(* IEC 61131-3 sources: 2026_Projet_YGO_ExcavatriceDragage/CODE_BACKUP/CODE_20260907_ChantierWeekEnd_v0.6.43/G_CYCLE/_TYPES, 10 files *)

(* ---- E_AutoCycleStep.st ---- *)
(* =======================================================================
   ⚙️ E_AutoCycleStep — Etapes du GRAFCET du cycle SEMI_AUTO (dragage)
   ───────────────────────────────────────────────────────────────
   🎯 Role : Enumeration des steps du sequenceur SEMI_AUTO (FB_CycleSemiAuto).
             Prefixe AX (Auto) homogene au homing machine (prefixe HX).
   📄 Doc metier : DOC/AF/AF_Partie-04_Mode_SemiAuto_Sequenceur_v2.3.md
                   + DOC/WFLOW/CONTRACTS/GEL_GRAFCET_SEMIAUTO_20260903.md
   🧊 GEL 2026-09-03 : DIVING decompose en 5 steps de plein droit (AX4..AX8) +
             step special AX_DIVING_RETRY ; EXTRACTION = AX9..AX12 ;
             DECHARGE = AX13..AX15C + AX18_DONE_SYNC ; AX_STAB repli defaut.
   ======================================================================= *)

TYPE E_AutoCycleStep :
(
  AX0_REPOS             := 0,   (* Repos / park : toutes commandes 0, etat neutre - etape initiale pure *)
  AX1_INIT             := 1,    (* Verif CONDITIONS INITIALES (Homed M1/M2, treuils FDC haut, M3 pas a droite de P1) - aucun mouvement, aucun referencement *)
  AX2_TRANSLATE_P1     := 2,    (* Translation vers P1 : joystick vers la droite, le cycle n'emet aucune commande M3 ; surveillance treuils au FDC haut *)
  AX3_OPEN_BUCKET      := 3,    (* Ouverture benne jusqu'au FDC logiciel benne ouverte *)

  (* --- DIVING (5 steps + retry) --- *)
  AX4_DESCEND_DIVING   := 4,    (* Plongee couplee benne ouverte palier 4 jusqu'a l'altimetrie de lancement (DiveStartMin_M) - Kobold PAS enclenche *)
  AX5_KOBOLD_INIT      := 5,    (* Activation contacteur Kobold << au vol >>, verif retour contacteur, descente palier 4 maintenue *)
  AX6_SEARCH_IMMERSION := 6,    (* Recherche entree dans l'eau : attente front DI Kobold 0->1, descente palier 4 maintenue *)
  AX7_SEARCH_BOTTOM    := 7,    (* Recherche du fond : attente front DI Kobold 1->0, descente palier 4 maintenue *)
  AX8_BOTTOM_CONFIRMED := 8,    (* Fond confirme : coupure instantanee treuils, set bit fond, TouchPositionM / RaiseTargetM *)

  (* --- EXTRACTION (4 steps) --- *)
  AX9_RAISE_OFF_BOTTOM := 9,    (* Montee synchronisee : retendre les cables ; selecteur couplage BOTH/M1/M2 accessible *)
  AX10_CLOSE_BUCKET    := 10,   (* Fermeture benne, treuils explicitement 0 *)
  AX11_CTRL_ASCENT     := 11,   (* Montee controle palier max reglable [1..2] + surveillance ecart vitesse M1/M2 ; benne mal fermee autorisee *)
  AX12_LOADED_ASCENT   := 12,   (* Montee en charge : palier 4 si benne fermee, palier 1 si mal fermee ; pas de ralenti 1 m avant top *)

  (* --- DECHARGE (6 steps) --- *)
  AX13_DRAIN_PAUSE     := 13,   (* Egouttage temporise - duree reglable IHM + bypass immediat *)
  AX14_TRANSLATE_DUMP  := 14,   (* Translation vers tremie (depart P1) + avertissements IHM *)
  AX15A_DUMP_ARRIVE    := 15,   (* Arrivee tremie : treuils a l'arret, attente geste operateur *)
  AX15B_DUMP_OPEN      := 16,   (* Vidage : ouverture benne au-dessus de la tremie, LES DEUX treuils a l'arret *)
  AX15C_DUMP_REPOSITION := 17,  (* Repositionnement couple M1+M2 (option IHM maintenue), retour AX15B au relachement *)
  AX18_DONE_SYNC       := 18,   (* Fin de passe : compteur vidages + duree cycle ; msg << aller en P1 >> ; rebouclage direct sur AX2 *)

  (* --- STEPS SPECIAUX --- *)
  AX_STAB              := 19,   (* Repli defaut / stabilisation - pas une erreur *)
  AX_DIVING_RETRY      := 20,   (* Reprise diving : remontee assistee palier lent jusqu'au FDC haut puis retour AX4 ; sur erreur Kobold / joystick relache / palier <> 4 en AX5..AX7 *)
  AX3_WAIT_DIVE_START  := 21,   (* Transition benne->plongee : sorties neutres jusqu'a l'arret mecanique confirme M1/M2, joystick pousse maintenu *)
  AX10_WAIT_ASCENT_START := 22  (* Transition fermeture->montee : sorties neutres jusqu'a l'arret confirme M1/M2, joystick tire maintenu *)
);
END_TYPE

(* ---- E_MachineHomingStep.st ---- *)
(* =======================================================================
   ⚙️ E_MachineHomingStep — Etapes du guide de referencement machine
   ───────────────────────────────────────────────────────────────
   🎯 Rôle : Etat publie du guide de homing conjoint M1/M2/benne (IHM + interlocks)
   📄 Doc métier : DOC/AF/AF_Partie-09_Fonction_Encoder_v2.4.md (F09.08)
   ======================================================================= *)

TYPE E_MachineHomingStep :
(
    IDLE                 := 0,   (* Referencement indisponible (Enable=FALSE) *)
    LOSS_SAFESTOP        := 5,   (* Perte de datum en mouvement : arret controle en cours *)
    BOTH_NOT_HOMED       := 10,  (* Codeurs M1 et M2 non references : passer en MAINT_N2 *)
    M1_NOT_HOMED         := 11,  (* Codeur M1 non reference ou mesure douteuse : homer M1 *)
    M2_NOT_HOMED         := 12,  (* Codeur M2 non reference ou mesure douteuse : homer M2 *)
    OFFSET_UNKNOWN       := 20,  (* Offset benne inconnu : passer en MAINT_N2 *)
    NEED_TOP_POSITION    := 30,  (* Monter Both a vitesse lente jusqu au capteur haut *)
    NEED_MECHANICAL_STOP := 40,  (* Capteur haut atteint : relacher la commande et attendre l arret *)
    AWAIT_BUCKET_CONFIRM := 45,  (* Confirmer visuellement la benne : Fermee ou Ouverte *)
    HOMING_IN_PROGRESS   := 50,  (* Referencement conjoint M1/M2 en cours : ne pas manoeuvrer *)
    VALID                := 60,  (* Referencement machine valide : mode nominal disponible *)
    FAILED               := 70   (* Referencement incomplet : rester en N2 et recommencer *)
);
END_TYPE

(* ---- E_MachineHomingTxState.st ---- *)
(* =======================================================================
   ⚙️ E_MachineHomingTxState — Steps du GRAFCET de referencement machine
   ───────────────────────────────────────────────────────────────
   🎯 Role : Machine a etats sequentielle (GRAFCET) du cycle de homing
             machine M1/M2/benne pilote par FB_CycleMachineHoming (§4).
             Distincte de E_MachineHomingStep (echelle de priorite du
             guide operateur, libelles de diagnostic - §6).
   📄 Doc : DOC/WFLOW/CONTRACTS/GEL_GRAFCET_HOMING_CYCLE_20260903.md
            + DOC/AF/AF_Partie-09_Fonction_Encoder_v2.4.md (F09.08)
   ======================================================================= *)

TYPE E_MachineHomingTxState :
(
    HX0_REPOS         := 0,   (* Etape initiale pure : aucune action, aucune affectation *)
    HX1_CHOICE        := 1,   (* Annonce + choix operateur : aucun mouvement *)
    HX2_CLIMB         := 2,   (* Chemin A : montee couplee M1+M2 palier 1 jusqu au capteur haut *)
    HX2N_NEUTRAL      := 3,   (* Arret + inversion de sens (tire -> pousse) : mouvement nul obligatoire *)
    HX3_HOME_AXES     := 4,   (* Homing axes M1+M2 au vol sur front descendant capteur, puis descente couplee *)
    HX3N_PAUSE        := 5,   (* Arret avant benne : mouvement nul, retour joystick au neutre *)
    HX4_BUCKET_ADJUST := 6,   (* Ajustement benne palier 1 sans FDC soft, 2 sens autorises *)
    HX5_BUCKET_COMMIT := 7,   (* Commit atomique etat benne fermee (CommitClose) *)
    HX6_HOMED         := 8,   (* Machine referencee : MachineHomed := TRUE (fugace) *)
    HXF_FAILED        := 9    (* Referencement incomplet : rester en N2 et recommencer *)
);
END_TYPE

(* ---- E_OperatorAxis.st ---- *)
(* =======================================================================
   ⚙️ E_OperatorAxis — Axe ou organe de pilotage attendu par le cycle
   ───────────────────────────────────────────────────────────────
   🎯 Rôle : Énumération de l'organe joystick/bouton attendu pour le mouvement
   📄 Doc métier : DOC/AF/AF_Partie-04_Mode_SemiAuto_Sequenceur_v2.3.md
   ======================================================================= *)

TYPE E_OperatorAxis :
(
    NONE        := 0, (* Aucun axe attendu (étape automatique ou arrêt) *)
    JOYSTICK_X  := 1, (* Axe X translation attendu *)
    JOYSTICK_Y  := 2, (* Axe Y treuils / plongée attendu *)
    BUTTON      := 3  (* Action bouton attendue (ex: validation, homing) *)
);
END_TYPE

(* ---- E_ProgramSequence.st ---- *)
(* =======================================================================
   ⚙️ E_ProgramSequence — Identifiant de la séquence programme active
   ───────────────────────────────────────────────────────────────
   🎯 Rôle : Identification de la séquence en cours d'exécution
   📄 Doc métier : DOC/AF/AF_Partie-04_Mode_SemiAuto_Sequenceur_v2.3.md
   ======================================================================= *)

TYPE E_ProgramSequence :
(
    NONE        := 0, (* Aucune séquence active *)
    MAIN_CYCLE  := 1, (* Cycle principal automatique de dragage X0..X13 *)
    DIVE_SEARCH := 2, (* Sous-séquence de plongée / recherche de fond *)
    EXTRACTION  := 3  (* Sous-séquence d'extraction et fermeture *)
);
END_TYPE

(* ---- ST_fbMachineHomingCycle_AxisHomingStatus.st ---- *)
(* =======================================================================
   🔌 ST_fbMachineHomingCycle_AxisHomingStatus — Statut homing d'un axe treuil
   ───────────────────────────────────────────────────────────────
   🎯 Rôle : Regroupe l'etat de homing d'un axe (M1 ou M2) consomme par
             FB_CycleMachineHoming pour piloter le guide et la transaction.
   📄 Doc métier : DOC/AF/AF_Partie-09_Fonction_Encoder_v2.4.md (F09.08)
   ======================================================================= *)
TYPE ST_fbMachineHomingCycle_AxisHomingStatus :
STRUCT
    HomedAndReliable : BOOL;   (* Codeur reference ET mesure jugee fiable (gate strict) *)
    HomingBusy       : BOOL;   (* Sequence de homing en cours sur l'axe *)
    HomingDone       : BOOL;   (* Homing termine avec succes (HomingLifecycle.Done cote FB_Encoder) *)
    HomingError      : BOOL;   (* Homing en erreur sur l'axe (HomingFault.Error) *)
END_STRUCT
END_TYPE

(* ---- ST_fbMachineHomingCycle_BucketCommit.st ---- *)
(* =======================================================================
   🔌 ST_fbMachineHomingCycle_BucketCommit — Commit atomique de l'etat benne
   ───────────────────────────────────────────────────────────────
   🎯 Rôle : Impulsion 1 scan emise par FB_CycleMachineHoming vers FB_Bucket
             apres succes des DEUX homings. FB_Bucket reste seul proprietaire
             de IsOpen / IsClosed.
   🔒 Sécurité : CommitOpen et CommitClose mutuellement exclusifs (garanti
                 par le corps du FB — rejet du double-confirm, cf. C-2).
   📄 Doc métier : DOC/AF/AF_Partie-05_Modes_Maintenance_v2.1.md
   ======================================================================= *)
TYPE ST_fbMachineHomingCycle_BucketCommit :
STRUCT
    CommitOpen  : BOOL;   (* Publier "benne ouverte" (impulsion 1 scan) *)
    CommitClose : BOOL;   (* Publier "benne fermee" (impulsion 1 scan) *)
END_STRUCT
END_TYPE

(* ---- ST_fbMachineHomingCycle_Cfg.st ---- *)
(* =======================================================================
   ⚙️ ST_fbMachineHomingCycle_Cfg — Réglages de FB_CycleMachineHoming
   ───────────────────────────────────────────────────────────────────────
   🎯 Rôle : Réglages géométriques du référencement machine (cible haute
             M2/benne + écarts benne) + temporisations de garde du GRAFCET
             de homing (montée, homing axes).
   🔒 Ownership : produit par PRG_02_Acquisition depuis _WinchM2CfgPersist
             (cible haute) et _BucketCfgPersist (écarts, GVL_PERSISTENT).
             Initialized : drapeau de restauration boot (pont persistant).
   📄 Doc métier : DOC/AF/AF_Partie-09_Fonction_Encoder_v2.4.md (F09.08)
   ======================================================================= *)

TYPE ST_fbMachineHomingCycle_Cfg :
STRUCT
    CfgTopHomingTarget_M : REAL;           // Position capteur haut M2/benne (m) — sert UNIQUEMENT a la cible dynamique M2 du cycle (HX3)
    CfgOffsetOpen_M      : REAL;           // Ecart géométrique benne ouverte (m)
    CfgOffsetClose_M     : REAL;           // Ecart géométrique benne fermée (m)
    CfgTimeoutClimb      : TIME := T#120s; // Garde HX2 : montée au capteur haut (0 = pas de garde)
    CfgTimeoutHomeAxes   : TIME := T#60s;  // Garde HX3 : descente jusqu'au front descendant capteur (0 = pas de garde)
    Initialized          : BOOL := FALSE;  // Drapeau de restauration config au boot (pont persistant)
END_STRUCT
END_TYPE

(* ---- ST_fbMachineHomingCycle_HomingDemand.st ---- *)
(* =======================================================================
   🔌 ST_fbMachineHomingCycle_HomingDemand — Demande de homing conjoint vers un axe
   ───────────────────────────────────────────────────────────────
   🎯 Rôle : Ordre de prise d'origine emis par FB_CycleMachineHoming vers
             une facade FB_Encoder. M1 : cible configuree. M2 : cible
             geometrique dynamique (top M1 configure +/- offset benne),
             jamais une position M1 live.
   📄 Doc métier : DOC/AF/AF_Partie-09_Fonction_Encoder_v2.4.md (F09.08)
   ======================================================================= *)
TYPE ST_fbMachineHomingCycle_HomingDemand :
STRUCT
    HomeReq          : BOOL;   (* Demande de prise d'origine pour cet axe (vocab reserve Homing) *)
    UseDynamicTarget : BOOL;   (* TRUE => cible = DynamicTarget_M (M2 uniquement) *)
    DynamicTarget_M  : REAL;   (* Cible geometrique benne (m) : CfgTopHomingTargetM + offset *)
END_STRUCT
END_TYPE

(* ---- ST_MachineHoming.st ---- *)
(* =======================================================================
   🧭 ST_MachineHoming — Etat publie du homing conjoint machine (M1/M2/benne)
   ───────────────────────────────────────────────────────────────
   🎯 Rôle : Regroupe les 8 sorties homing a plat de PRG_02_Acquisition en
             un bus struct unique, publie sur le bus inter-PRG.
   🔒 Sécurité : Homed = qualification conjointe reference machine (gate SEMI_AUTO).
                 HomingLoss = perte reference en mouvement : arret controle SafeStop.
   📄 Doc métier : DOC/AF/AF_Partie-09_Fonction_Encoder_v2.4.md (F09.08)
   ======================================================================= *)
TYPE ST_MachineHoming :
STRUCT
    Homed            : BOOL;          (* Qualification conjointe reference machine *)
    SetPosBucketOpen : BOOL;          (* Valider position actuelle = reference benne ouverte *)
    SetPosBucketClose: BOOL;          (* Valider position actuelle = reference benne fermee *)
    Active           : BOOL;          (* Homing conjoint en cours *)
    HomingLoss       : BOOL;          (* Perte reference en mouvement : arret controle SafeStop *)
    Step             : INT;           (* Etape guidee reference (echelle de priorite E_MachineHomingStep) *)
    Instruction      : STRING(120);   (* Consigne IHM reference *)
    Failed           : BOOL;          (* Transaction reference abandonnee *)
    SeqStep          : INT;           (* Step GRAFCET courant (E_MachineHomingTxState HX0..HXF) *)
    M3Locked         : BOOL;          (* Translation M3 interdite pendant le cycle de homing machine *)
    CmdWinchM1       : ST_ProgramWinchRequest; (* Ordre treuil M1 couple palier 1 (HX2 montee / HX3 descente) *)
    CmdWinchM2       : ST_ProgramWinchRequest; (* Ordre treuil M2 couple palier 1 (HX2 montee / HX3 descente) *)
    CmdBucketOpen    : BOOL;          (* Ordre ouverture benne palier 1 sans FDC soft (HX4) *)
    CmdBucketClose   : BOOL;          (* Ordre fermeture benne palier 1 sans FDC soft (HX4) *)
END_STRUCT
END_TYPE
